// TIA Portal V20 export
Screen "StyleOverview"  1276x673
  ScreenItem "Title_OPMode1_ScreenOverview_X390_Y2" at 493,7 size 500x30  Type=HmiTextBox
  ScreenItem "Button_Back" at 11,0 size 117x42  Type=HmiButton
  ScreenItem "Button_26" at 0,0 size 126x22  Type=HmiButton
  ScreenItem "Button_7" at 0,22 size 126x19  Type=HmiButton
  ScreenItem "Button_2" at 0,41 size 126x19  Type=HmiButton
  ScreenItem "Button_1" at 0,60 size 126x19  Type=HmiButton
  ScreenItem "Button_4" at 0,79 size 126x19  Type=HmiButton
  ScreenItem "Button_6" at 0,118 size 126x19  Type=HmiButton
  ScreenItem "Button_8" at 0,136 size 126x23  Type=HmiButton
  ScreenItem "Button_9" at 0,159 size 126x19  Type=HmiButton
  ScreenItem "Button_24" at 0,98 size 126x20  Type=HmiButton
  ScreenItem "Button_31" at 0,176 size 126x23  Type=HmiButton
  ScreenItem "Button_17" at 0,0 size 126x22  Type=HmiButton
  ScreenItem "Button_16" at 0,22 size 126x19  Type=HmiButton
  ScreenItem "Button_15" at 0,41 size 126x19  Type=HmiButton
  ScreenItem "Button_14" at 0,60 size 126x19  Type=HmiButton
  ScreenItem "Button_13" at 0,79 size 126x19  Type=HmiButton
  ScreenItem "Button_11" at 0,118 size 126x19  Type=HmiButton
  ScreenItem "Button_10" at 0,136 size 126x23  Type=HmiButton
  ScreenItem "Button_5" at 0,159 size 126x19  Type=HmiButton
  ScreenItem "Button_12" at 0,98 size 126x20  Type=HmiButton
  ScreenItem "Button_3" at 0,176 size 126x23  Type=HmiButton
  ScreenItem "Button_40" at 0,0 size 126x22  Type=HmiButton
  ScreenItem "Button_39" at 0,22 size 126x19  Type=HmiButton
  ScreenItem "Button_38" at 0,41 size 126x19  Type=HmiButton
  ScreenItem "Button_37" at 0,60 size 126x19  Type=HmiButton
  ScreenItem "Button_36" at 0,79 size 126x19  Type=HmiButton
  ScreenItem "Button_34" at 0,118 size 126x19  Type=HmiButton
  ScreenItem "Button_33" at 0,136 size 126x23  Type=HmiButton
  ScreenItem "Button_32" at 0,159 size 126x19  Type=HmiButton
  ScreenItem "Button_35" at 0,98 size 126x20  Type=HmiButton
  ScreenItem "Button_30" at 0,176 size 126x23  Type=HmiButton
  ScreenItem "面板容器_8" at 151,40 size 204x210  Type=HmiFaceplateContainer
  ScreenItem "面板容器_9" at 377,40 size 204x210  Type=HmiFaceplateContainer
  ScreenItem "面板容器_3" at 603,40 size 204x210  Type=HmiFaceplateContainer
  ScreenItem "面板容器_16" at 829,40 size 204x210  Type=HmiFaceplateContainer
  ScreenItem "面板容器_5" at 1055,40 size 204x216  Type=HmiFaceplateContainer
  ScreenItem "面板容器_1" at 151,246 size 204x210  Type=HmiFaceplateContainer
  ScreenItem "面板容器_2" at 377,246 size 204x210  Type=HmiFaceplateContainer
  ScreenItem "面板容器_6" at 603,246 size 204x210  Type=HmiFaceplateContainer
  ScreenItem "面板容器_7" at 829,246 size 204x210  Type=HmiFaceplateContainer
  ScreenItem "面板容器_10" at 1055,246 size 204x210  Type=HmiFaceplateContainer
  ScreenItem "Button_20" at 0,0 size 126x22  Type=HmiButton
  ScreenItem "Button_18" at 0,22 size 126x19  Type=HmiButton
  ScreenItem "Button_19" at 0,41 size 126x19  Type=HmiButton
  ScreenItem "Button_28" at 0,60 size 126x19  Type=HmiButton
  ScreenItem "Button_21" at 0,79 size 126x19  Type=HmiButton
  ScreenItem "Button_23" at 0,118 size 126x19  Type=HmiButton
  ScreenItem "Button_25" at 0,136 size 126x23  Type=HmiButton
  ScreenItem "Button_27" at 0,159 size 126x19  Type=HmiButton
  ScreenItem "Button_22" at 0,98 size 126x20  Type=HmiButton
  ScreenItem "Button_29" at 0,176 size 126x23  Type=HmiButton
  ScreenItem "面板容器_4" at 151,452 size 204x210  Type=HmiFaceplateContainer
  ScreenItem "面板容器_11" at 377,452 size 204x210  Type=HmiFaceplateContainer
  ScreenItem "面板容器_12" at 603,452 size 204x210  Type=HmiFaceplateContainer
  ScreenItem "面板容器_13" at 829,452 size 204x210  Type=HmiFaceplateContainer
